(* IEC 61131-3 sources: codesys-api/examples/mqtt_large_payload/st, 4 files *)

(* ---- AppendText.st ---- *)
FUNCTION AppendText : BOOL
// Appends Text to a long STRING without CONCAT, which stops at 255 characters.
// Returns FALSE and leaves the buffer unchanged when Text would not fit.
VAR_INPUT
	pBuffer : POINTER TO BYTE;  // ADR() of the destination STRING
	Capacity : UDINT;           // SIZEOF() of the destination, terminator included
	Text : STRING(255);         // one short piece; only the total may exceed 255
END_VAR
VAR_IN_OUT
	Used : UDINT;               // current length of the destination, kept by the caller
END_VAR
VAR
	pText : POINTER TO BYTE;
	TextLength : UDINT;
	Index : UDINT;
END_VAR
// ---- implementation ----
TextLength := INT_TO_UDINT(LEN(Text));
IF pBuffer = 0 OR Used + TextLength + 1 > Capacity THEN
	AppendText := FALSE;
	RETURN;
END_IF

pText := ADR(Text);
FOR Index := 1 TO TextLength DO
	pBuffer[Used] := pText[Index - 1];
	Used := Used + 1;
END_FOR
pBuffer[Used] := 0;
AppendText := TRUE;

(* ---- NowUs.st ---- *)
FUNCTION NowUs : ULINT
// Monotonic microsecond clock for the performance counters.
VAR
	Microseconds : ULINT;
END_VAR
// ---- implementation ----
SysTimeCore.SysTimeGetUs(pUsTime := Microseconds);
NowUs := Microseconds;

(* ---- PLC_PRG.BuildLine.st ---- *)
// Action BuildLine: sets Line to payload line number Index (0-based), newline included.
// Value i is Sequence*1000 + i, or that divided by 100 as a two-decimal REAL.
// ---- implementation ----
IF Index = 0 THEN
	Line := CONCAT('DEMO_SEQ:', UDINT_TO_STRING(Sequence));
ELSIF Index = 1 THEN
	Line := CONCAT('DEMO_COUNT:', UINT_TO_STRING(ValueCount));
ELSIF Index = 2 THEN
	Line := SEL(IsRealFormat, 'DEMO_FORMAT:INT', 'DEMO_FORMAT:REAL');
ELSIF Index = ValueCount + 3 THEN
	Line := CONCAT('DEMO_END:', UDINT_TO_STRING(Sequence));
ELSE
	ValueIndex := Index - 2;
	Line := CONCAT(CONCAT('DEMO_V', UINT_TO_STRING(ValueIndex)), ':');
	IF IsRealFormat THEN
		RealValue := UDINT_TO_REAL(Sequence * 1000 + UINT_TO_UDINT(ValueIndex)) / 100.0;
		// The same rounding and conversion as BCNF's FB_InterlockMatrix.StringPublication.
		Line := CONCAT(Line, REAL_TO_STRING(DINT_TO_REAL(TRUNC(RealValue * 100.0 + SEL(RealValue >= 0.0, -0.5, 0.5))) / 100.0));
	ELSE
		Line := CONCAT(Line, UDINT_TO_STRING(Sequence * 1000 + UINT_TO_UDINT(ValueIndex)));
	END_IF
END_IF
Line := CONCAT(Line, '$N');

(* ---- PLC_PRG.st ---- *)
PROGRAM PLC_PRG
// Publishes one large MQTT payload with the unmodified Stefan Dreyer MQTT 1.2.0.7 library.
// Optionally also publishes a CONCAT-built copy of the same text, which shows where the
// 255-character cap comes from; it is off by default so the timings match production.
// The *Us/*Cycles variables measure what large payloads cost the PLC; write ResetStats to clear maxima.
VAR
	MqttLink : MQTT.MQTT_IN_OUT;          // not "Mqtt": ST names are case-insensitive and would hide the MQTT namespace
	LargePublisher : MQTT.MQTTPublish;
	ConcatPublisher : MQTT.MQTTPublish;
	IsInitialized : BOOL;

	// Settings, writable online
	BrokerUrl : STRING(250) := '192.168.50.240:1883';
	LargeTopic : STRING(64) := 'raw_data_demo';
	ConcatTopic : STRING(64) := 'raw_data_demo/concat';
	ValueCount : UINT := 500;            // values per message
	PublishPeriod : TIME := T#1S;        // BCNF publishes once a second
	IsRealFormat : BOOL := TRUE;         // two-decimal REALs formatted the way BCNF does; FALSE = integers
	IsQos1 : BOOL := FALSE;              // BCNF publishes at QoS 0
	IsConcatControlEnabled : BOOL;       // the 255-character demonstration; not production work
	IsBcnfEveryScanEnabled : BOOL;       // run BCNF's StringPublication (verbatim copy) every scan, as BCNF does
	IsTagValueEnabled : BOOL;            // publish BCNF's values as tag:value lines once a second
	TagValueTopic : STRING(64) := 'raw_data_demo/tagvalue';
	ClientCallsPerScan : INT := 1;       // most client calls per scan while a message is in flight (one 4 KB buffer per two calls)
	ClientBudgetUs : ULINT := 5000;      // ... and stop calling once this much time went into the client this scan
	IsClientLoopGated : BOOL := TRUE;    // FALSE: always make ClientCallsPerScan calls (to measure idle calls)
	ClientSlots : UINT := 40;            // out slots of the MQTT client (library default 16; recommended 8, here 40
	                                     // so SplitTest can keep 32 messages in flight)
	ClientSlotsIn : UINT := 20;          // in slots. mochi sends QoS 1/2 without an inflight limit; a QoS 2 burst with more
	                                     // messages than this and over 16 KB waits on PUBRELs it cannot read (disconnect)

	IsClientCalledLast : BOOL;           // run the client loop at the end of the scan, after the publishers
	IsSecondClientCallEnabled : BOOL;    // call the client once more at the end of the scan, after the publishers,
	                                     // so a reply requested in this scan goes out in this scan (latency test)
	IsSendInFlight : BOOL;
	ClientCall : INT;
	MaxClientCalls : INT;
	IsCopyBenchRequested : BOOL;         // time the library's payload copy: MEM.MemMove of one 4,095-byte send buffer
	CopyBuffer : ARRAY[0..4095] OF BYTE;
	CopyBenchUs : UDINT;                 // mean of 20 copies
	PublishTimer : TON;

	LargePayload : STRING(30000);        // about 1,500 two-decimal values
	LargeUsed : UDINT;
	ConcatPayload : STRING(8000);        // the "bigger string" approach that still truncates
	Line : STRING(80);                   // one short line; CONCAT is fine below 255
	PublishQoS : MQTT.QoS;

	IsLargeRequested : BOOL;
	IsConcatRequested : BOOL;
	IsBuildOk : BOOL;
	Sequence : UDINT;
	Index : UINT;
	ValueIndex : UINT;
	RealValue : REAL;

	// Diagnostics, readable online
	IsBrokerConnected : BOOL;
	LargeSentCount : UDINT;
	ConcatSentCount : UDINT;
	TimeoutCount : UDINT;
	OverflowCount : UDINT;
	SkippedBusyCount : UDINT;
	LastLargeLength : UDINT;
	LastConcatLength : UDINT;

	// Performance, microseconds unless named *Cycles
	ResetStats : BOOL;
	CycleStartUs : ULINT;
	PreviousCycleStartUs : ULINT;
	StepStartUs : ULINT;
	LargeRequestUs : ULINT;
	LastLargeBuildUs : UDINT;
	MaxLargeBuildUs : UDINT;
	LastConcatBuildUs : UDINT;
	MaxConcatBuildUs : UDINT;
	ClientUs : UDINT;
	MaxClientUs : UDINT;
	SecondCallBudgetUs : UDINT := 2000;  // the second call runs only if the first took less than this
	SecondStartUs : ULINT;
	SecondClientUs : UDINT;
	ScanClientUs : UDINT;                // both calls in this scan
	MaxScanClientUs : UDINT;
	CycleUs : UDINT;
	MaxCycleUs : UDINT;
	IntervalUs : UDINT;
	MaxIntervalUs : UDINT;
	MinIntervalUs : UDINT := 16#FFFFFFFF;
	LargeBusyCycles : UDINT;
	LastPublishCycles : UDINT;
	MaxPublishCycles : UDINT;
	LastPublishUs : UDINT;
	MaxPublishUs : UDINT;
	LastBcnfBuildUs : UDINT;             // one call of BCNF's StringPublication copy
	MaxBcnfBuildUs : UDINT;
	BcnfBuildCount : UDINT;
	BcnfBuildTotalUs : ULINT;            // average = BcnfBuildTotalUs / BcnfBuildCount

	// BCNF's values in tag:value format (BcnfStringPublicationCopy.BuildTagValue), built once per publish
	TagValuePublisher : MQTT.MQTTPublish;
	TagValueTimer : TON;
	TagValueQoS : MQTT.QoS;
	IsTagValueRequested : BOOL;
	TagValueRequestUs : ULINT;
	TagValueBusyCycles : UDINT;
	TagValueSentCount : UDINT;
	TagValueTimeoutCount : UDINT;
	LastTagValueLength : UDINT;
	LastTagValueBuildUs : UDINT;
	MaxTagValueBuildUs : UDINT;
	TagValueBuildCount : UDINT;
	TagValueBuildTotalUs : ULINT;
	LastTagValuePublishUs : UDINT;
	MaxTagValuePublishUs : UDINT;
	LastTagValuePublishCycles : UDINT;
	MaxTagValuePublishCycles : UDINT;
END_VAR
// ---- implementation ----
CycleStartUs := NowUs();
IF IsCopyBenchRequested THEN
	IsCopyBenchRequested := FALSE;
	StepStartUs := NowUs();
	FOR Index := 1 TO 20 DO
		MEM.MemMove(pSource := ADR(LargePayload), pDestination := ADR(CopyBuffer), uiNumberOfBytes := 4095);
	END_FOR
	CopyBenchUs := ULINT_TO_UDINT(NowUs() - StepStartUs) / 20;
END_IF

IF ResetStats THEN
	ResetStats := FALSE;
	MaxLargeBuildUs := 0;
	MaxConcatBuildUs := 0;
	MaxClientUs := 0;
	MaxScanClientUs := 0;
	MaxClientCalls := 0;
	MaxCycleUs := 0;
	MaxIntervalUs := 0;
	MinIntervalUs := 16#FFFFFFFF;
	MaxPublishCycles := 0;
	MaxPublishUs := 0;
	PreviousCycleStartUs := 0;
	MaxBcnfBuildUs := 0;
	BcnfBuildCount := 0;
	BcnfBuildTotalUs := 0;
	MaxTagValueBuildUs := 0;
	TagValueBuildCount := 0;
	TagValueBuildTotalUs := 0;
	MaxTagValuePublishUs := 0;
	MaxTagValuePublishCycles := 0;
END_IF
IF PreviousCycleStartUs <> 0 THEN
	IntervalUs := ULINT_TO_UDINT(CycleStartUs - PreviousCycleStartUs);
	MaxIntervalUs := MAX(MaxIntervalUs, IntervalUs);
	MinIntervalUs := MIN(MinIntervalUs, IntervalUs);
END_IF
PreviousCycleStartUs := CycleStartUs;

MqttLink.ClientID := 'BENCH_MQTT_DEMO';
// Incoming publishes up to 40 KB of payload (EdgeTest); the library's default limit is 2,000 bytes of payload
// plus the largest topic. Read once, at the client's first call.
MqttLink.COM_CONFIG.MaxPayloadSize := 40000;
// Slots for messages in flight; the library walks every slot on every call. The demo has six publishers and
// one subscriber; the library default is 50 each way. Read once, at the client's first call.
MqttLink.COM_CONFIG.CountSlotsIn := ClientSlotsIn;
MqttLink.COM_CONFIG.CountSlotsOut := ClientSlots;
// The client moves one 4 KB send buffer per two calls. While any message is in flight, call it again until
// ClientCallsPerScan calls or ClientBudgetUs; otherwise once, for keep-alive and receiving.
IF NOT IsClientCalledLast THEN
	CallClient();
END_IF
IsBrokerConnected := MqttLink.BROKER_CONNECTED;

IF NOT IsInitialized THEN
	IsInitialized := TRUE;
	LargePublisher.SetMqttInOut(MQTT_IN_OUT := MqttLink);
	ConcatPublisher.SetMqttInOut(MQTT_IN_OUT := MqttLink);
	TagValuePublisher.SetMqttInOut(MQTT_IN_OUT := MqttLink);
END_IF

PublishTimer(IN := NOT PublishTimer.Q, PT := PublishPeriod);

// The library reads the payload through its pointer over several cycles,
// so a payload is only rebuilt once its previous publish has finished.
IF PublishTimer.Q AND IsBrokerConnected THEN
	IF IsLargeRequested OR IsConcatRequested THEN
		SkippedBusyCount := SkippedBusyCount + 1;
	ELSE
		Sequence := Sequence + 1;
		// Lines: DEMO_SEQ, DEMO_COUNT, DEMO_FORMAT, DEMO_V1..DEMO_Vn, DEMO_END (see BuildLine).
		StepStartUs := NowUs();
		LargeUsed := 0;
		LargePayload := '';
		IsBuildOk := TRUE;
		FOR Index := 0 TO ValueCount + 3 DO
			BuildLine();
			IsBuildOk := IsBuildOk AND AppendText(pBuffer := ADR(LargePayload), Capacity := SIZEOF(LargePayload), Text := Line, Used := LargeUsed);
		END_FOR
		LastLargeBuildUs := ULINT_TO_UDINT(NowUs() - StepStartUs);
		MaxLargeBuildUs := MAX(MaxLargeBuildUs, LastLargeBuildUs);

		ConcatPayload := '';
		LastConcatBuildUs := 0;
		IF IsConcatControlEnabled THEN
			StepStartUs := NowUs();
			FOR Index := 0 TO ValueCount + 3 DO
				BuildLine();
				ConcatPayload := CONCAT(ConcatPayload, Line);
			END_FOR
			LastConcatBuildUs := ULINT_TO_UDINT(NowUs() - StepStartUs);
			MaxConcatBuildUs := MAX(MaxConcatBuildUs, LastConcatBuildUs);
		END_IF

		IF NOT IsBuildOk THEN
			OverflowCount := OverflowCount + 1;
		END_IF
		LastLargeLength := LargeUsed;
		LastConcatLength := INT_TO_UDINT(LEN(ConcatPayload));
		IF IsQos1 THEN
			PublishQoS := MQTT.QoS.AtLeastOnce;
		ELSE
			PublishQoS := MQTT.QoS.AtMostOnce;
		END_IF
		IsLargeRequested := IsBuildOk;
		IsConcatRequested := IsConcatControlEnabled;
		LargeRequestUs := NowUs();
		LargeBusyCycles := 0;
	END_IF
END_IF

LargePublisher(
	Topic := ADR(LargeTopic),
	PayloadString := ADR(LargePayload),
	PublishAsString := TRUE,
	QoSIn := PublishQoS,
	MRetain := FALSE,
	send := IsLargeRequested);

ConcatPublisher(
	Topic := ADR(ConcatTopic),
	PayloadString := ADR(ConcatPayload),
	PublishAsString := TRUE,
	QoSIn := PublishQoS,
	MRetain := FALSE,
	send := IsConcatRequested AND NOT IsLargeRequested);

IF IsLargeRequested THEN
	LargeBusyCycles := LargeBusyCycles + 1;
END_IF
IF LargePublisher.done THEN
	IsLargeRequested := FALSE;
	LargeSentCount := LargeSentCount + 1;
	// Request to done: PUBACK at QoS 1, payload handed to TCP at QoS 0; includes the scans spent copying it out.
	LastPublishUs := ULINT_TO_UDINT(NowUs() - LargeRequestUs);
	MaxPublishUs := MAX(MaxPublishUs, LastPublishUs);
	LastPublishCycles := LargeBusyCycles;
	MaxPublishCycles := MAX(MaxPublishCycles, LastPublishCycles);
END_IF
IF ConcatPublisher.done THEN
	IsConcatRequested := FALSE;
	ConcatSentCount := ConcatSentCount + 1;
END_IF
IF LargePublisher.SendTimeout OR ConcatPublisher.SendTimeout THEN
	TimeoutCount := TimeoutCount + 1;
	IsLargeRequested := FALSE;
	IsConcatRequested := FALSE;
END_IF

// BCNF's values as tag:value lines: built only in the scan that publishes, sent as one message.
IF IsQos1 THEN
	TagValueQoS := MQTT.QoS.AtLeastOnce;
ELSE
	TagValueQoS := MQTT.QoS.AtMostOnce;
END_IF
TagValueTimer(IN := IsTagValueEnabled AND NOT TagValueTimer.Q, PT := T#1S);
IF TagValueTimer.Q AND IsBrokerConnected AND NOT IsTagValueRequested THEN
	StepStartUs := NowUs();
	BcnfStringPublicationCopy.BuildTagValue();
	LastTagValueBuildUs := ULINT_TO_UDINT(NowUs() - StepStartUs);
	MaxTagValueBuildUs := MAX(MaxTagValueBuildUs, LastTagValueBuildUs);
	TagValueBuildCount := TagValueBuildCount + 1;
	TagValueBuildTotalUs := TagValueBuildTotalUs + LastTagValueBuildUs;
	LastTagValueLength := BcnfStringPublicationCopy.TagValueUsed;
	IsTagValueRequested := BcnfStringPublicationCopy.IsTagValueBuildOk;
	TagValueRequestUs := NowUs();
	TagValueBusyCycles := 0;
END_IF
TagValuePublisher(
	Topic := ADR(TagValueTopic),
	PayloadString := ADR(BcnfStringPublicationCopy.TagValuePayload),
	PublishAsString := TRUE,
	QoSIn := TagValueQoS,
	MRetain := FALSE,
	send := IsTagValueRequested);
IF IsTagValueRequested THEN
	TagValueBusyCycles := TagValueBusyCycles + 1;
END_IF
IF TagValuePublisher.done THEN
	IsTagValueRequested := FALSE;
	TagValueSentCount := TagValueSentCount + 1;
	LastTagValuePublishUs := ULINT_TO_UDINT(NowUs() - TagValueRequestUs);
	MaxTagValuePublishUs := MAX(MaxTagValuePublishUs, LastTagValuePublishUs);
	LastTagValuePublishCycles := TagValueBusyCycles;
	MaxTagValuePublishCycles := MAX(MaxTagValuePublishCycles, LastTagValuePublishCycles);
END_IF
IF TagValuePublisher.SendTimeout THEN
	TagValueTimeoutCount := TagValueTimeoutCount + 1;
	IsTagValueRequested := FALSE;
END_IF

// UTC from the NTP server for the scale test's timestamps (and the PLC's clock, if enabled).
ClockSync();

// 2,000-tag scale test (idle unless ScaleTest.IsEnabled); inside the timed scan on purpose.
ScaleTest();
// MQTT library edge-case test (idle unless EdgeTest.IsEnabled; edge_test.py drives it).
EdgeTest();
// The same data as one message or many (idle unless SplitTest.IsEnabled; split_test.py drives it).
SplitTest();
// Mixed-rate load: 75 % of the tags once a second, 25 % ten times a second (idle unless MixedTest.IsEnabled; mixed_rate_test.py).
MixedTest();
// BCNF's own MQTT code with its two client connections (idle unless BcnfComms.IsEnabled; bcnf_test.py drives it).
BcnfComms();
// Rewritten by online_change_test.py to make online changes (does nothing else).
OnlineChangeProbe();
// Broker URL parsing check (idle unless UrlProbe.Input is written; url_test.py).
UrlProbe();
// The second call sends what the publishers requested in this scan (a command's acknowledgement), but only
// while the first call left room in the scan's client budget: during a full refresh the first call already
// sent a 16 KB buffer, and a second one would double the scan's client time.
SecondClientUs := 0;
IF IsSecondClientCallEnabled AND ClientUs < SecondCallBudgetUs THEN
	SecondStartUs := NowUs();
	MqttLink.clientFB(MQTT_IN_OUT := MqttLink, ENABLE := TRUE, URL := BrokerUrl, TIMEOUT := T#10S, TLS := FALSE);
	SecondClientUs := ULINT_TO_UDINT(NowUs() - SecondStartUs);
END_IF
ScanClientUs := ClientUs + SecondClientUs;
MaxScanClientUs := MAX(MaxScanClientUs, ScanClientUs);
// With IsClientCalledLast the client runs once per scan here, after every publisher and subscriber, so a
// reply requested in this scan goes out in this scan's call.
IF IsClientCalledLast THEN
	CallClient();
END_IF

// What BCNF pays today: its payload strings are rebuilt in every scan, not only when publishing.
IF IsBcnfEveryScanEnabled THEN
	StepStartUs := NowUs();
	BcnfStringPublicationCopy();
	LastBcnfBuildUs := ULINT_TO_UDINT(NowUs() - StepStartUs);
	MaxBcnfBuildUs := MAX(MaxBcnfBuildUs, LastBcnfBuildUs);
	BcnfBuildCount := BcnfBuildCount + 1;
	BcnfBuildTotalUs := BcnfBuildTotalUs + LastBcnfBuildUs;
END_IF

CycleUs := ULINT_TO_UDINT(NowUs() - CycleStartUs);
MaxCycleUs := MAX(MaxCycleUs, CycleUs);
